FUNCTION_BLOCK logiBUS_QD_PWM (* Output service interface function block for 13-bit PWM output data (0..8191 in DWORD) *)
  (* Description: Copyright (c) 2017 fortiss GmbH, HR Agrartechnik GmbH This program and the accompanying materials are made available under the terms of the Eclipse Public License 2.0 which is available at https://www.eclipse.org/legal/epl-2.0/ SPDX-License-Identifier: EPL-2.0 *)
  (* Version 1.2, 2026-11-06, Franz Höpfinger, Meisterschulen am Ostbahnhof, Add FREQ, RAMP and RAMPO (hardware ramp, LEDC timer pool) *)
  (* Version 1.1, 2026-09-20, Franz Höpfinger, Meisterschulen am Ostbahnhof, Document 13-bit resolution (0..8191, 0..100% duty cycle) for OUT variable *)
  (* Version 1.0, 2017-03-20, Monika Wenger, fortiss GmbH, initial API and implementation and/or initial documentation *)
  PACKAGE logiBUS::io::DQ;
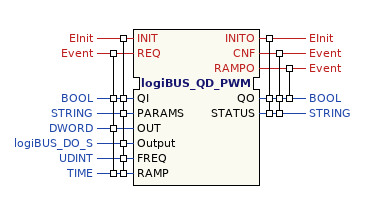
  EVENT_INPUT
    INIT : EInit WITH QI, PARAMS, Output, FREQ, RAMP; (* Service Initialization *)
    REQ WITH QI, OUT, RAMP; (* Service Request *)
  END_EVENT
  EVENT_OUTPUT
    INITO : EInit WITH QO, STATUS; (* Initialization Confirm *)
    CNF WITH QO, STATUS; (* Confirmation of Requested Service *)
    RAMPO WITH QO; (* Ramp finished: OUT reached (immediately after the jump with RAMP = T#0ms) *)
  END_EVENT
  VAR_INPUT
    QI : BOOL; (* Event Input Qualifier *)
    PARAMS : STRING; (* Service Parameters *)
    OUT : DWORD; (* 13-bit raw PWM output value (0..8191, 0..100% duty cycle) *)
    Output : logiBUS::io::DQ::logiBUS_DO_S := logiBUS_DO::Invalid; (* Identify the Output Output_Q1..Q8 *)
    FREQ : UDINT := 400; (* PWM frequency in Hz, read at INIT. Outputs with the same frequency share an LEDC timer (4 timers, LED blinking uses one). Power stage limits, not checked: APIXON 15 PWR Q1 (BTH50030) max. 100 Hz; BTS7030/BTT6030/BTH6070 for valves 100..200 Hz; Trainer20 without power stage *)
    RAMP : TIME := T#0ms; (* Transition time to the new OUT value (hardware ramp), read at INIT and REQ. T#0ms = jump *)
  END_VAR
  VAR_OUTPUT
    QO : BOOL; (* Event Output Qualifier *)
    STATUS : STRING; (* Service Status *)
  END_VAR
END_FUNCTION_BLOCK
